(* IEC 61131-3 sources: codesys-to-s7/tests/corpus/C2S7-TYPE-64/pos, 1 file *)

(* ---- input.st ---- *)
FUNCTION_BLOCK FB_Case
VAR
    q : LINT;
END_VAR
q := 1;
END_FUNCTION_BLOCK
